Staubli VAL3: getCurMoveID.pgx

public program getCurMoveID(bool x_bGetMoveId, string x_sType)
  local bool l_bGetMoveId
begin
  l_bGetMoveId=(x_bGetMoveId==true)
  if !l_bGetMoveId
    if(x_sType=="Stop" or x_sType=="Abort" or x_sType=="End") and !bHaveGetMoveID
      nCurrentMoveID=getMoveId()
      bHaveGetMoveID=true
    endIf
    // bInterrupt=true
  else
    bInterrupt=true
  endIf
end
